{attribute 'qualified_only'}
{attribute 'strict'}
TYPE E_CIP_Source :
(
	eNone := 0,
	eT91_Sanitation,
	eT92_Detergent,
	eT93_R_Water,
	eT94_Water,
	eClose
);
END_TYPE

(* stored: Version 1.1.0.1, ProductVersion 3.1.4024.12
   DUT E_CIP_Source: Id {0e935b9e-07f5-4e10-94ab-b8db9546b09f} *)
